{attribute 'pack_mode' := '1'}
TYPE ST_ScheduleWork_V1 :
STRUCT
 DeviceID : UDINT;
 WeekDay : UDINT;
 StartTime : UINT;
 EndTime : UINT;
 Value : REAL;
 Operation : UDINT;
END_STRUCT
END_TYPE

(* stored: Version 1.1.0.1, ProductVersion 3.1.4024.15
   DUT ST_ScheduleWork_V1: Id {4463d85b-444f-4689-9986-49d67fcaf9c2} *)
